    dio dDio = {link=0AE8B5A8-7356-480B-AAA1-20AFD496F398}
    string sComment = "备用"
  [125]
    dio dDio = {link=DB043A0E-80EF-4F10-9CBC-7A049A7AEFDE}
    string sComment = "备用"
  [126]
    dio dDio = {link=951CF18F-CA29-47EF-A085-39A8D6CD28C1}
    string sComment = "备用"
  [127]
    dio dDio = {link=6FC2F7D5-08CF-47CC-86FA-1AC31B966FFD}
    string sComment = "备用"
public dioItem dOutItem[128]
  [0]
    dio dDio = {link=813E3F4B-A1DE-4C5D-8EAB-0242B6D8A546}
    string sComment = "外部内模式"
  [1]
    dio dDio = {link=364EC08F-C077-495B-A954-158507D3C26C}
    string sComment = "机器人上电状态"
  [2]
    dio dDio = {link=289A5E8D-11F3-4BEB-8FA4-200735E3A2B7}
    string sComment = "程序运行中"
  [3]
    dio dDio = {link=79705501-C546-4790-A460-3F340ADFDE5C}
    string sComment = "机器人报警"
  [4]
    dio dDio = {link=75D4F3C1-C356-4EDA-B423-02C90835EA7D}
    string sComment = "机器人急停"
  [5]
    dio dDio = {link=3F319035-E82A-4D07-9742-3AFC501B53DF}
    string sComment = "备用"
  [6]
    dio dDio = {link=1CC4B59E-3D71-495F-A34B-473B0A37D044}
    string sComment = "备用"
  [7]
    dio dDio = {link=2087A18A-21B3-4E9A-90F0-0A72D013BBC2}
    string sComment = "备用"
  [8]
    dio dDio = {link=93BF17B5-5C7E-43C6-9C42-3B6025772815}
    string sComment = "机器人作业原点"
  [9]
    dio dDio = {link=16CB4CF9-3A13-4F09-B6E9-D967DFB15E25}
    string sComment = "机器人喷涂中"
  [10]
    dio dDio = {link=734EBAF3-2CA8-4D3F-A8BB-E168C1322725}
    string sComment = "机器人开关枪"
  [11]
    dio dDio = {link=07A4EEA8-4CAE-47C3-9487-42EFEC0C0C8E}
    string sComment = "喷涂完成"
  [12]
    dio dDio = {link=63159677-63A9-4936-A8C6-E65B2885D59F}
    string sComment = "备用"
  [13]
    dio dDio = {link=698A0489-9B90-43A7-B0CD-777095A36007}
    string sComment = "备用"
  [14]
    dio dDio = {link=C4522756-21A9-4D8A-B398-209F6EFB0977}
    string sComment = "备用"
  [15]
    dio dDio = {link=E3974102-9CCD-497B-BD29-7D9DDF1F0662}
    string sComment = "备用"
  [16]
    dio dDio = {link=D7E9BDA6-AD73-4469-BD4D-C9D8F1711105}
    string sComment = "备用"
  [17]
    dio dDio = {link=C0E9CDD3-3C86-4E8A-BB76-29DD4E724269}
    string sComment = "备用"
  [18]
    dio dDio = {link=19A15CFF-CD59-4687-8101-878C6D297AD0}
    string sComment = "备用"
  [19]
    dio dDio = {link=F886CB4C-7C2D-4AEE-8DA8-19CCB8826A1C}
    string sComment = "备用"
  [20]
    dio dDio = {link=44B2E852-2BDD-46AD-B032-142EDC75806B}
    string sComment = "备用"
  [21]
    dio dDio = {link=E6202C42-8108-4A9C-988A-BA326395584A}
    string sComment = "备用"
  [22]
    dio dDio = {link=4A293BE2-BE94-462E-ACFA-7E01BA496DDB}
    string sComment = "备用"
  [23]
    dio dDio = {link=C4CC4269-4D2F-4B53-89D1-5B6F0F9E20C5}
    string sComment = "备用"
  [24]
    dio dDio = {link=976E4904-0F44-43DA-867D-0C06FC7F067A}
    string sComment = "备用"
  [25]
    dio dDio = {link=26F2F168-65FE-450B-BE6F-27BCBE8A7C37}
    string sComment = "备用"
  [26]
    dio dDio = {link=58979B7C-3302-40C0-9293-D8BDE318359F}
    string sComment = "备用"
  [27]
    dio dDio = {link=32E62FFE-3CE0-449B-8ADB-B460A9E5DE54}
    string sComment = "备用"
  [28]
    dio dDio = {link=1778E8D0-D57F-4F6E-A6A4-A7E0DC8A5FDF}
    string sComment = "备用"
  [29]
    dio dDio = {link=BB6EEE31-C681-41BA-8160-A41199CEAD02}
    string sComment = "备用"
  [30]
    dio dDio = {link=58577585-C0FF-479D-B4D2-FF8F04E87201}
    string sComment = "备用"
  [31]
    dio dDio = {link=E4789C35-874D-4E09-8AF9-741C03AAD9B4}
    string sComment = "备用"
  [32]
    dio dDio = {link=AB4C11BC-0698-4F05-9F77-33C54B19FD7D}
    string sComment = "备用"
  [33]
    dio dDio = {link=A971CAAA-D369-4C08-BB4B-F444CDC4D2F0}
    string sComment = "备用"
  [34]
    dio dDio = {link=EE574E0A-35B5-4DE1-8C9E-C0DF9CDCDFE6}
    string sComment = "备用"
  [35]
    dio dDio = {link=7532402E-1B90-4BA9-83CA-579B1F726874}
    string sComment = "备用"
  [36]
    dio dDio = {link=6F6C7C8F-8851-47C2-9B8E-D33C24B9D39F}
    string sComment = "备用"
  [37]
    dio dDio = {link=4A5CAAE4-C9CD-4421-94AD-56079246CA39}
    string sComment = "备用"
  [38]
    dio dDio = {link=EB7E2C34-F887-4C3F-97E0-01834D630C5E}
    string sComment = "备用"
  [39]
    dio dDio = {link=BDBB409A-6EC7-4423-9FF9-A638D02BF80E}
    string sComment = "备用"
  [40]
    dio dDio = {link=E136414E-B9B9-4DA1-8541-C1A78F1E80BF}
    string sComment = "备用"
  [41]
    dio dDio = {link=8E4798E6-5BA8-40FC-8B4C-D83695D2AB51}
    string sComment = "备用"
  [42]
    dio dDio = {link=28472F68-DF34-4C50-9023-A219CE2C4B1B}
    string sComment = "备用"
  [43]
    dio dDio = {link=1DB5BD39-DE07-40ED-B700-8C7874B04DB0}
    string sComment = "备用"
  [44]
    dio dDio = {link=88484DFD-5685-4FE3-BD11-1467A80C9B34}
    string sComment = "备用"
  [45]
    dio dDio = {link=2F5F1623-83AA-4A31-A803-F6FA4D4BE14A}
    string sComment = "备用"
  [46]
    dio dDio = {link=519B5132-0D61-4FA5-ABD4-96724AED25E8}
    string sComment = "备用"
  [47]
    dio dDio = {link=661BE778-7099-413C-A47D-EC9A4ECEF23E}
    string sComment = "备用"
  [48]
    dio dDio = {link=53B2124C-FE98-440B-9A3D-84530B55B740}
    string sComment = "备用"
  [49]
    dio dDio = {link=229E980F-A7B4-4859-9EE1-BA541F4B5A16}
    string sComment = "备用"
  [50]
    dio dDio = {link=1FA4F26D-23CC-42E9-A819-02B2DD7006DA}
    string sComment = "备用"
  [51]
    dio dDio = {link=2AEDD394-CA8D-4F24-A299-43D2A058ACD5}
    string sComment = "备用"
  [52]
    dio dDio = {link=C28EB1DF-BACA-4254-A598-B532E330438E}
    string sComment = "备用"
  [53]
    dio dDio = {link=E7F3183B-4DF3-459A-ADF7-79D82988755C}
    string sComment = "备用"
  [54]
    dio dDio = {link=2614E536-799A-40AF-9560-80A760021F62}
    string sComment = "备用"
  [55]
    dio dDio = {link=757B7056-4991-459D-8227-2BCDF4BE047B}
    string sComment = "备用"
  [56]
    dio dDio = {link=8C99F1DA-9DA9-4BDF-B60F-FD54ABC54EFA}
    string sComment = "备用"
  [57]
    dio dDio = {link=5AA809C1-68E1-4A24-9F04-C8074121C64A}
    string sComment = "备用"
  [58]
    dio dDio = {link=4A164529-4FC6-4374-9AB6-7CFCFB13974B}
    string sComment = "备用"
  [59]
    dio dDio = {link=70724C45-B1FB-42FE-A3A2-C0AB8AA81684}
    string sComment = "备用"
  [60]
    dio dDio = {link=9EE71F53-97CD-4882-A49E-A6F1E8BC9441}
    string sComment = "4ST总工位完成"
  [61]
    dio dDio = {link=81277848-FDAC-47B2-B4F0-EFE16B2F5C1C}
    string sComment = "第1步；4ST-紊流清洗1  完成"
  [62]
    dio dDio = {link=E56352E6-5F75-449C-AD2C-249D38B077FB}
    string sComment = "第2步；4ST机器人工作1   完成"
  [63]
    dio dDio = {link=5728C013-0742-4355-8E61-1A03F1F076E6}
    string sComment = "第3步；4ST-翻转180清洗15S  完成"
  [64]
    dio dDio = {link=04B33B81-599B-4BDE-99DF-EEC79DF42297}
    string sComment = "第4步；4ST-紊流清洗1(5度25)   完成"
  [65]
    dio dDio = {link=D5C4F9D4-602E-45CC-A360-A9C8DFC51706}
    string sComment = "第5步；4ST  控水：180：30S//-180：30S 完成"
  [66]
    dio dDio = {link=0F23F4DE-A6DC-48A8-BD13-38096E17E4BC}
    string sComment = "第6步；4ST机器人工作:吹干 完成"
  [67]
    dio dDio = {link=725D593E-3E8C-49B9-A0C8-EC5E7EDBEF47}
    string sComment = "第7步；4ST  控水：180：30S//-180：30S 完成"
  [68]
    dio dDio = {link=D80F8BA0-A9D7-467A-84F3-2EF911086F28}
    string sComment = "备用"
  [69]
    dio dDio = {link=290333BB-E8D8-473B-B7DA-1770BF97A3BA}
    string sComment = "备用"
  [70]
    dio dDio = {link=3451ABCB-1CE5-49F5-8053-7E43529834C5}
    string sComment = "备用"
  [71]
    dio dDio = {link=1C486D5A-1AEA-494E-AC84-6CEA9FC0F052}
    string sComment = "备用"
  [72]
    dio dDio = {link=0B5202A6-62EE-4D6C-8E76-4A396B266DA1}
    string sComment = "备用"
  [73]
    dio dDio = {link=07376469-6AEC-4E90-A30D-02A336A51CCF}
    string sComment = "备用"
  [74]
    dio dDio = {link=9C60D734-A29B-44DA-837E-97A014720D64}
    string sComment = "备用"
  [75]
    dio dDio = {link=F6F5CEBA-7A13-4322-B86E-E02B17A52B8C}
    string sComment = "备用"
  [76]
    dio dDio = {link=034F848A-A2B4-4107-BA29-37F2DF0B4836}
    string sComment = "备用"
  [77]
    dio dDio = {link=2D3AB11E-A0E7-43D6-A64B-B19DE4EDCA54}
    string sComment = "备用"
  [78]
    dio dDio = {link=6B87E34F-9D7F-4178-ADAD-CF451768FAD1}
    string sComment = "备用"
  [79]
    dio dDio = {link=0BECC0A6-11C6-443C-B8B7-B823C5449F03}
    string sComment = "备用"
  [80]
    dio dDio = {link=0FAFA963-6C61-46BA-8B8E-FD5D821CED0B}
    string sComment = "备用"
  [81]
    dio dDio = {link=E858B3E5-8FFB-4B3B-9E73-58A45F891801}
    string sComment = "备用"
  [82]
    dio dDio = {link=52490A38-A31A-4D56-AA93-4E3292557F7F}
    string sComment = "备用"
  [83]
    dio dDio = {link=07DE5AAD-9C80-4970-8E40-B99AD098B2C3}
    string sComment = "备用"
  [84]
    dio dDio = {link=E76E3858-8352-4107-BC87-39491D8B651A}
    string sComment = "备用"
  [85]
    dio dDio = {link=2B09FA37-BF2E-4ED9-B53F-09BB42630F57}
    string sComment = "备用"
  [86]
    dio dDio = {link=C0D4BCE7-AA67-4991-AD3B-5583CCFF9A80}
    string sComment = "备用"
  [87]
    dio dDio = {link=BBA329F0-9B99-401C-B2C0-5AA54B82A434}
    string sComment = "备用"
  [88]
    dio dDio = {link=1FF771B4-EE27-450D-A9DB-7E394712BF39}
    string sComment = "备用"
  [89]
    dio dDio = {link=19978664-DA67-4FAE-9478-F6C2FD7BC1A1}
    string sComment = "备用"
  [90]
    dio dDio = {link=B280086E-4E78-4C33-A16A-5103EDFD12BA}
    string sComment = "备用"
  [91]
    dio dDio = {link=66D76411-AF4D-465C-BF45-D26D600CE49D}
    string sComment = "备用"
  [92]
    dio dDio = {link=CF5BF486-B482-4F9A-936E-D7550E22D48F}
    string sComment = "备用"
  [93]
    dio dDio = {link=47EF2689-3337-4012-BAD2-52612379B15C}
    string sComment = "备用"
  [94]
    dio dDio = {link=9BC9630D-0782-4292-B056-6CBDA421EF62}
    string sComment = "备用"
  [95]
    dio dDio = {link=CAFB5CCA-B450-480D-9CAD-A29B903F45A9}
    string sComment = "备用"
  [96]
    dio dDio = {link=DCBA4C7F-A728-4F25-89A5-B6259619A80B}
    string sComment = "参考位置1"
  [97]
    dio dDio = {link=6753AC4A-51FA-413E-B4B2-137174F0D507}
    string sComment = "参考位置2"
  [98]
    dio dDio = {link=81370562-9275-47C1-93C0-CB31297CDD20}
    string sComment = "参考位置3"
  [99]
    dio dDio = {link=E6DCC6F0-C964-47CD-B4D7-1BD8BFDA33AE}
    string sComment = "参考位置4"
  [100]
    dio dDio = {link=18C334B4-AE06-448E-96BF-3CD280A2541B}
    string sComment = "参考位置5"
  [101]
    dio dDio = {link=15B48D0D-C668-47AF-A704-10BA0ED6FFE7}
    string sComment = "参考位置6"
  [102]
    dio dDio = {link=DA2930BB-B07C-4C38-ADBB-0FDC55ECF2BB}
    string sComment = "参考位置7"
  [103]
    dio dDio = {link=8DDD8F2E-B5A8-4F54-BD1B-48D04A96C878}
    string sComment = "参考位置8"
  [104]
    dio dDio = {link=72245E17-FF99-4704-8474-EDB79B027BF9}
    string sComment = "参考位置9"
  [105]
    dio dDio = {link=BCF85E34-592F-4BA5-AE76-F1E8F2FD96C1}
    string sComment = "参考位置10"
  [106]
    dio dDio = {link=9ED9CFBB-1644-41A9-955E-D6E7EB6EF2F1}
    string sComment = "参考位置11"
  [107]
    dio dDio = {link=5A6FDD52-29C6-40B7-B97D-88DE84ED4E53}
    string sComment = "参考位置12"
  [108]
    dio dDio = {link=8E4836F5-8A3D-4937-90E9-0F98CBF16A27}
    string sComment = "参考位置13"
  [109]
    dio dDio = {link=4305B788-10E3-4C38-9835-3E94A9820D41}
    string sComment = "参考位置14"
  [110]
    dio dDio = {link=152B6212-6AC5-4D19-A5F9-C32452DCD0BD}
    string sComment = "参考位置15"
  [111]
    dio dDio = {link=60BD22D0-03A0-4632-85E7-7AB9A7B5E9EE}
    string sComment = "参考位置16"
  [112]
    dio dDio = {link=617AC81D-63D2-418A-A221-1A45E82E8F33}
    string sComment = "干涉区1"
  [113]
    dio dDio = {link=DA60158B-5C4B-4C1D-9AEB-3A4C25735862}
    string sComment = "干涉区2"
  [114]
    dio dDio = {link=7E45E59A-6E5F-4DD8-8E87-A62787B5121D}
    string sComment = "干涉区3"
  [115]
    dio dDio = {link=302676B4-AFEF-4A5D-9D0F-7D7EEE15BD09}
    string sComment = "干涉区4"
  [116]
    dio dDio = {link=94FD2E61-B0C4-426E-8CB5-3D13DE4E72D1}
    string sComment = "干涉区5"
  [117]
    dio dDio = {link=5441B2EB-7737-420D-A838-CB6BC6A9AA98}
    string sComment = "干涉区6"
  [118]
    dio dDio = {link=D70A9639-74F8-485B-B1AE-A12B6619BE09}
    string sComment = "干涉区7"
  [119]
    dio dDio = {link=3C4D5DF3-3DD0-4928-9BAC-FF9DB40E9304}
    string sComment = "干涉区8"
  [120]
    dio dDio = {link=389B2383-01D9-4D6D-8093-13CF39736E4D}
    string sComment = "干涉区9"
  [121]
    dio dDio = {link=9C61CF1A-5A0B-480F-A9AF-E365017F4409}
    string sComment = "干涉区10"
  [122]
    dio dDio = {link=D6F4FFC6-5A52-44AE-AAFC-981F5DBD7076}
    string sComment = "干涉区11"
  [123]
    dio dDio = {link=3768B870-3C40-471D-B639-CE39EBCB3865}
    string sComment = "干涉区12"
  [124]
    dio dDio = {link=FCBA4290-2AF9-4EDB-AAB3-C3D5B2BC56ED}
    string sComment = "干涉区13"
  [125]
    dio dDio = {link=FEB8E5C1-4C55-454A-AACA-1D927BE28924}
    string sComment = "干涉区14"
  [126]
    dio dDio = {link=C97B50B1-B825-4E71-A20E-3BFEC37BB4DF}
    string sComment = "干涉区15"
  [127]
    dio dDio = {link=FB88829F-F043-4942-9C93-D2BA50858194}
    string sComment = "干涉区16"
public num nMaxAnalog = 8
public num nMaxdigital = 128
public num nProgfb
public string sCommentAin[24]
  [0] = "接收程序号"
  [1] = "刷子号反馈"
  [2] = "备用"
  [3] = "备用"
  [4] = "备用"
  [5] = "备用"
  [6] = "备用"
  [7] = "备用"
  [8] = "备用"
  [9] = "备用"
  [10] = "备用"
  [11] = "备用"
  [12] = "备用"
  [13] = "备用"
  [14] = "备用"
  [15] = "备用"
  [16] = "备用"
  [17] = "备用"
  [18] = "备用"
  [19] = "备用"
  [20] = "备用"
  [21] = "备用"
  [22] = "备用"
  [23] = "备用"
public string sCommentAout[24]
  [0] = "程序号反馈"
  [1] = "刷子号"
  [2] = "备用"
  [3] = "备用"
  [4] = "备用"
  [5] = "备用"
  [6] = "备用"
  [7] = "备用"
  [8] = "备用"
  [9] = "备用"
  [10] = "备用"
  [11] = "备用"
  [12] = "备用"
  [13] = "备用"
  [14] = "备用"
  [15] = "备用"
  [16] = "备用"
  [17] = "备用"
  [18] = "备用"
  [19] = "备用"
  [20] = "备用"
  [21] = "备用"
  [22] = "备用"
  [23] = "备用"
public string sCommentDin[128]
  [0] = "电机上电"
  [1] = "主程序运行"
  [2] = "复位报警"
  [3] = "PLC系统故障"
  [4] = "备用"
  [5] = "备用"
  [6] = "备用"
  [7] = "备用"
  [8] = "开枪完成"
  [9] = "关枪完成"
  [10] = "开始喷涂"
  [11] = "备用"
  [12] = "备用"
  [13] = "备用"
  [14] = "备用"
  [15] = "备用"
  [16] = "备用"
  [17] = "备用"
  [18] = "备用"
  [19] = "备用"
  [20] = "备用"
  [21] = "备用"
  [22] = "备用"
  [23] = "备用"
  [24] = "备用"
  [25] = "备用"
  [26] = "备用"
  [27] = "备用"
  [28] = "备用"
  [29] = "备用"
  [30] = "备用"
  [31] = "备用"
  [32] = "备用"
  [33] = "备用"
  [34] = "备用"
  [35] = "备用"
  [36] = "备用"
  [37] = "备用"
  [38] = "备用"
  [39] = "备用"
  [40] = "备用"
  [41] = "备用"
  [42] = "备用"
  [43] = "备用"
  [44] = "备用"
  [45] = "备用"
  [46] = "备用"
  [47] = "备用"
  [48] = "备用"
  [49] = "备用"
  [50] = "备用"
  [51] = "备用"
  [52] = "备用"
  [53] = "备用"
  [54] = "备用"
  [55] = "备用"
  [56] = "备用"
  [57] = "备用"
  [58] = "备用"
  [59] = "备用"
  [60] = "备用"
  [61] = "备用"
  [62] = "备用"
  [63] = "备用"
  [64] = "备用"
  [65] = "备用"
  [66] = "备用"
  [67] = "备用"
  [68] = "备用"
  [69] = "备用"
  [70] = "备用"
  [71] = "备用"
  [72] = "备用"
  [73] = "备用"
  [74] = "备用"
  [75] = "备用"
  [76] = "备用"
  [77] = "备用"
  [78] = "备用"
  [79] = "备用"
  [80] = "备用"
  [81] = "备用"
  [82] = "备用"
  [83] = "备用"
  [84] = "备用"
  [85] = "备用"
  [86] = "备用"
  [87] = "备用"
  [88] = "备用"
  [89] = "备用"
  [90] = "备用"
  [91] = "备用"
  [92] = "备用"
  [93] = "备用"
  [94] = "备用"
  [95] = "备用"
  [96] = "备用"
  [97] = "备用"
  [98] = "备用"
  [99] = "备用"
  [100] = "备用"
  [101] = "备用"
  [102] = "备用"
  [103] = "备用"
  [104] = "备用"
  [105] = "备用"
  [106] = "备用"
  [107] = "备用"
  [108] = "备用"
  [109] = "备用"
  [110] = "备用"
  [111] = "备用"
  [112] = "备用"
  [113] = "备用"
  [114] = "备用"
  [115] = "备用"
  [116] = "备用"
  [117] = "备用"
  [118] = "备用"
  [119] = "备用"
  [120] = "备用"
  [121] = "备用"
  [122] = "备用"
  [123] = "备用"
  [124] = "备用"
  [125] = "备用"
  [126] = "备用"
  [127] = "备用"
public string sCommentDout[128]
  [0] = "外部内模式"
  [1] = "机器人上电状态"
  [2] = "程序运行中"
  [3] = "机器人报警"
  [4] = "机器人急停"
  [5] = "备用"
  [6] = "备用"
  [7] = "备用"
  [8] = "机器人作业原点"
  [9] = "机器人喷涂中"
  [10] = "机器人开关枪"
  [11] = "喷涂完成"
  [12] = "备用"
  [13] = "备用"
  [14] = "备用"
  [15] = "备用"
  [16] = "备用"
  [17] = "备用"
  [18] = "备用"
  [19] = "备用"
  [20] = "备用"
  [21] = "备用"
  [22] = "备用"
  [23] = "备用"
  [24] = "备用"
  [25] = "备用"
  [26] = "备用"
  [27] = "备用"
  [28] = "备用"
  [29] = "备用"
  [30] = "备用"
  [31] = "备用"
  [32] = "备用"
  [33] = "备用"
  [34] = "备用"
  [35] = "备用"
  [36] = "备用"
  [37] = "备用"
  [38] = "备用"
  [39] = "备用"
  [40] = "备用"
  [41] = "备用"
  [42] = "备用"
  [43] = "备用"
  [44] = "备用"
  [45] = "备用"
  [46] = "备用"
  [47] = "备用"
  [48] = "备用"
  [49] = "备用"
  [50] = "备用"
  [51] = "备用"
  [52] = "备用"
  [53] = "备用"
  [54] = "备用"
  [55] = "备用"
  [56] = "备用"
  [57] = "备用"
  [58] = "备用"
  [59] = "备用"
  [60] = "4ST总工位完成"
  [61] = "第1步；4ST-紊流清洗1  完成"
  [62] = "第2步；4ST机器人工作1   完成"
  [63] = "第3步；4ST-翻转180清洗15S  完成"
  [64] = "第4步；4ST-紊流清洗1(5度25)   完成"
  [65] = "第5步；4ST  控水：180：30S//-180：30S 完成"
  [66] = "第6步；4ST机器人工作:吹干 完成"
  [67] = "第7步；4ST  控水：180：30S//-180：30S 完成"
  [68] = "备用"
  [69] = "备用"
  [70] = "备用"
  [71] = "备用"
  [72] = "备用"
  [73] = "备用"
  [74] = "备用"
  [75] = "备用"
  [76] = "备用"
  [77] = "备用"
  [78] = "备用"
  [79] = "备用"
  [80] = "备用"
  [81] = "备用"
  [82] = "备用"
  [83] = "备用"
  [84] = "备用"
  [85] = "备用"
  [86] = "备用"
  [87] = "备用"
  [88] = "备用"
  [89] = "备用"
  [90] = "备用"
  [91] = "备用"
  [92] = "备用"
  [93] = "备用"
  [94] = "备用"
  [95] = "备用"
  [96] = "参考位置1"
  [97] = "参考位置2"
  [98] = "参考位置3"
  [99] = "参考位置4"
  [100] = "参考位置5"
  [101] = "参考位置6"
  [102] = "参考位置7"
  [103] = "参考位置8"
  [104] = "参考位置9"
  [105] = "参考位置10"
  [106] = "参考位置11"
  [107] = "参考位置12"
  [108] = "参考位置13"
  [109] = "参考位置14"
  [110] = "参考位置15"
  [111] = "参考位置16"
  [112] = "干涉区1"
  [113] = "干涉区2"
  [114] = "干涉区3"
  [115] = "干涉区4"
  [116] = "干涉区5"
  [117] = "干涉区6"
  [118] = "干涉区7"
  [119] = "干涉区8"
  [120] = "干涉区9"
  [121] = "干涉区10"
  [122] = "干涉区11"
  [123] = "干涉区12"
  [124] = "干涉区13"
  [125] = "干涉区14"
  [126] = "干涉区15"
  [127] = "干涉区16"
